                                           #StatConfigDigital[#temp16IndexDigital].OSLevel := #ConfigDint[#temp16IndexDigital].OSLevel;
                                           #StatConfigDigital[#temp16IndexDigital].ApplyExt := #ConfigDint[#temp16IndexDigital].ApplyExt;
                                           #StatConfigDigital[#temp16IndexDigital].ApplyOp := #ConfigDint[#temp16IndexDigital].ApplyOp;
                                           #StatConfigDigital[#temp16IndexDigital].Sync := #ConfigDint[#temp16IndexDigital].Sync;
                                           #StatConfigDigital[#temp16IndexDigital].StateOffOp := #ConfigDint[#temp16IndexDigital].StateOffOp;
                                           #StatConfigDigital[#temp16IndexDigital].StateOpOp := #ConfigDint[#temp16IndexDigital].StateOpOp;
                                           #StatConfigDigital[#temp16IndexDigital].StateAutOp := #ConfigDint[#temp16IndexDigital].StateAutOp;
                                           #StatConfigDigital[#temp16IndexDigital].SrcIntOp := #ConfigDint[#temp16IndexDigital].SrcIntOp;
                                           #StatConfigDigital[#temp16IndexDigital].SrcExtOp := #ConfigDint[#temp16IndexDigital].SrcExtOp;
                                           #StatConfigDigital[#temp16IndexDigital].VExt := #ConfigDint[#temp16IndexDigital].VExt;
                                           #StatConfigDigital[#temp16IndexDigital].VOp := #ConfigDint[#temp16IndexDigital].VOp;
                                       END_IF;
                                       #temp16IndexDigital := #temp16IndexDigital + 1;
                                   END_REGION
                                   // If Parameter type = 3(Binary)
                               #TYPE_BINARY:
                                   REGION Binary
                                       //Bit Masking funtionality for calculate the used Binary parameter
                                       #ConfigParaType.IndexBinary := #ConfigParaType.IndexBinary OR SHL(IN := #temp32TempDword1, N := INT_TO_UINT(#temp16IndexOfDefinition));
                                       //Condition to check the config binary parameters are within range 
                                       IF ((#temp16IndexIO >= #CONFIG_PARAMETER_MIN) AND (#temp16IndexIO <= #MAPPED_CONFIG_BINARY)) THEN
                                           //WinCC Parameter View Faceplate logic
                                           #ConfigBin[#temp16IndexBinary].WQC := #ConfigurationParameterBinary[#temp16IndexMTP].WQC;
                                           #ConfigBin[#temp16IndexBinary].ApplyEn := #ConfigurationParameterBinary[#temp16IndexMTP].ApplyEn;
                                           #ConfigBin[#temp16IndexBinary].ApplyInt := #ConfigurationParameterBinary[#temp16IndexMTP].ApplyInt;
                                           #ConfigBin[#temp16IndexBinary].StateChannel := #ConfigurationParameterBinary[#temp16IndexMTP].StateChannel;
                                           #ConfigBin[#temp16IndexBinary].StateOffAut := #ConfigurationParameterBinary[#temp16IndexMTP].StateOffAut;
                                           #ConfigBin[#temp16IndexBinary].StateOpAut := #ConfigurationParameterBinary[#temp16IndexMTP].StateOpAut;
                                           #ConfigBin[#temp16IndexBinary].StateAutAut := #ConfigurationParameterBinary[#temp16IndexMTP].StateAutAut;
                                           #ConfigBin[#temp16IndexBinary].StateOffAct := #ConfigurationParameterBinary[#temp16IndexMTP].StateOffAct;
                                           #ConfigBin[#temp16IndexBinary].StateOpAct := #ConfigurationParameterBinary[#temp16IndexMTP].StateOpAct;
                                           #ConfigBin[#temp16IndexBinary].StateAutAct := #ConfigurationParameterBinary[#temp16IndexMTP].StateAutAct;
                                           #ConfigBin[#temp16IndexBinary].SrcChannel := #ConfigurationParameterBinary[#temp16IndexMTP].SrcChannel;
                                           #ConfigBin[#temp16IndexBinary].SrcExtAut := #ConfigurationParameterBinary[#temp16IndexMTP].SrcExtAut;
                                           #ConfigBin[#temp16IndexBinary].SrcIntAut := #ConfigurationParameterBinary[#temp16IndexMTP].SrcIntAut;
                                           #ConfigBin[#temp16IndexBinary].SrcIntAct := #ConfigurationParameterBinary[#temp16IndexMTP].SrcIntAct;
                                           #ConfigBin[#temp16IndexBinary].SrcExtAct := #ConfigurationParameterBinary[#temp16IndexMTP].SrcExtAct;
                                           #ConfigBin[#temp16IndexBinary].VInt := #ConfigurationParameterBinary[#temp16IndexMTP].VInt;
                                           #ConfigBin[#temp16IndexBinary].VReq := #ConfigurationParameterBinary[#temp16IndexMTP].VReq;
                                           #ConfigBin[#temp16IndexBinary].VOut := #ConfigurationParameterBinary[#temp16IndexMTP].VOut;
                                           #ConfigBin[#temp16IndexBinary].VFbk := #ConfigurationParameterBinary[#temp16IndexMTP].VFbk;
                                           #ConfigBin[#temp16IndexBinary].VState0 := #ConfigurationParameterBinary[#temp16IndexMTP].VState0;
                                           #ConfigBin[#temp16IndexBinary].VState1 := #ConfigurationParameterBinary[#temp16IndexMTP].VState1;
                                           //Write values from WinCC
                                           IF #ConfigurationParameterBinary[#temp16IndexMTP].OSLevel = #StatConfigBinary[#temp16IndexBinary].OSLevel THEN
                                               #ConfigurationParameterBinary[#temp16IndexMTP].OSLevel := #ConfigBin[#temp16IndexBinary].OSLevel;
                                           ELSE
                                               #ConfigBin[#temp16IndexBinary].OSLevel := #ConfigurationParameterBinary[#temp16IndexMTP].OSLevel;
                                           END_IF;
                                           IF #ConfigurationParameterBinary[#temp16IndexMTP].ApplyExt = #StatConfigBinary[#temp16IndexBinary].ApplyExt THEN
                                               #ConfigurationParameterBinary[#temp16IndexMTP].ApplyExt := #ConfigBin[#temp16IndexBinary].ApplyExt;
                                           ELSE
                                               #ConfigBin[#temp16IndexBinary].ApplyExt := #ConfigurationParameterBinary[#temp16IndexMTP].ApplyExt;
                                           END_IF;
                                           IF #ConfigurationParameterBinary[#temp16IndexMTP].ApplyOp = #StatConfigBinary[#temp16IndexBinary].ApplyOp THEN
                                               #ConfigurationParameterBinary[#temp16IndexMTP].ApplyOp := #ConfigBin[#temp16IndexBinary].ApplyOp;
                                           ELSE
                                               #ConfigBin[#temp16IndexBinary].ApplyOp := #ConfigurationParameterBinary[#temp16IndexMTP].ApplyOp;
                                           END_IF;
                                           IF #ConfigurationParameterBinary[#temp16IndexMTP].Sync = #StatConfigBinary[#temp16IndexBinary].Sync THEN
                                               #ConfigurationParameterBinary[#temp16IndexMTP].Sync := #ConfigBin[#temp16IndexBinary].Sync;
                                           ELSE
                                               #ConfigBin[#temp16IndexBinary].Sync := #ConfigurationParameterBinary[#temp16IndexMTP].Sync;
                                           END_IF;
                                           IF #ConfigurationParameterBinary[#temp16IndexMTP].StateOffOp = #StatConfigBinary[#temp16IndexBinary].StateOffOp THEN
                                               #ConfigurationParameterBinary[#temp16IndexMTP].StateOffOp := #ConfigBin[#temp16IndexBinary].StateOffOp;
                                           ELSE
                                               #ConfigBin[#temp16IndexBinary].StateOffOp := #ConfigurationParameterBinary[#temp16IndexMTP].StateOffOp;
                                           END_IF;
                                           IF #ConfigurationParameterBinary[#temp16IndexMTP].StateOpOp = #StatConfigBinary[#temp16IndexBinary].StateOpOp THEN
                                               #ConfigurationParameterBinary[#temp16IndexMTP].StateOpOp := #ConfigBin[#temp16IndexBinary].StateOpOp;
                                           ELSE
                                               #ConfigBin[#temp16IndexBinary].StateOpOp := #ConfigurationParameterBinary[#temp16IndexMTP].StateOpOp;
                                           END_IF;
                                           IF #ConfigurationParameterBinary[#temp16IndexMTP].StateAutOp = #StatConfigBinary[#temp16IndexBinary].StateAutOp THEN
                                               #ConfigurationParameterBinary[#temp16IndexMTP].StateAutOp := #ConfigBin[#temp16IndexBinary].StateAutOp;
                                           ELSE
                                               #ConfigBin[#temp16IndexBinary].StateAutOp := #ConfigurationParameterBinary[#temp16IndexMTP].StateAutOp;
                                           END_IF;
                                           IF #ConfigurationParameterBinary[#temp16IndexMTP].SrcIntOp = #StatConfigBinary[#temp16IndexBinary].SrcIntOp THEN
                                               #ConfigurationParameterBinary[#temp16IndexMTP].SrcIntOp := #ConfigBin[#temp16IndexBinary].SrcIntOp;
                                           ELSE
                                               #ConfigBin[#temp16IndexBinary].SrcIntOp := #ConfigurationParameterBinary[#temp16IndexMTP].SrcIntOp;
                                           END_IF;
                                           IF #ConfigurationParameterBinary[#temp16IndexMTP].SrcExtOp = #StatConfigBinary[#temp16IndexBinary].SrcExtOp THEN
                                               #ConfigurationParameterBinary[#temp16IndexMTP].SrcExtOp := #ConfigBin[#temp16IndexBinary].SrcExtOp;
                                           ELSE
                                               #ConfigBin[#temp16IndexBinary].SrcExtOp := #ConfigurationParameterBinary[#temp16IndexMTP].SrcExtOp;
                                           END_IF;
                                           IF #ConfigurationParameterBinary[#temp16IndexMTP].VExt = #StatConfigBinary[#temp16IndexBinary].VExt THEN
                                               #ConfigurationParameterBinary[#temp16IndexMTP].VExt := #ConfigBin[#temp16IndexBinary].VExt;
                                           ELSE
                                               #ConfigBin[#temp16IndexBinary].VExt := #ConfigurationParameterBinary[#temp16IndexMTP].VExt;
                                           END_IF;
                                           IF #ConfigurationParameterBinary[#temp16IndexMTP].VOp = #StatConfigBinary[#temp16IndexBinary].VOp THEN
                                               #ConfigurationParameterBinary[#temp16IndexMTP].VOp := #ConfigBin[#temp16IndexBinary].VOp;
                                           ELSE
                                               #ConfigBin[#temp16IndexBinary].VOp := #ConfigurationParameterBinary[#temp16IndexMTP].VOp;
                                           END_IF;

                                           #StatConfigBinary[#temp16IndexBinary].OSLevel := #ConfigBin[#temp16IndexBinary].OSLevel;
                                           #StatConfigBinary[#temp16IndexBinary].ApplyExt := #ConfigBin[#temp16IndexBinary].ApplyExt;
                                           #StatConfigBinary[#temp16IndexBinary].ApplyOp := #ConfigBin[#temp16IndexBinary].ApplyOp;
                                           #StatConfigBinary[#temp16IndexBinary].Sync := #ConfigBin[#temp16IndexBinary].Sync;
                                           #StatConfigBinary[#temp16IndexBinary].StateOffOp := #ConfigBin[#temp16IndexBinary].StateOffOp;
                                           #StatConfigBinary[#temp16IndexBinary].StateOpOp := #ConfigBin[#temp16IndexBinary].StateOpOp;
                                           #StatConfigBinary[#temp16IndexBinary].StateAutOp := #ConfigBin[#temp16IndexBinary].StateAutOp;
                                           #StatConfigBinary[#temp16IndexBinary].SrcIntOp := #ConfigBin[#temp16IndexBinary].SrcIntOp;
                                           #StatConfigBinary[#temp16IndexBinary].SrcExtOp := #ConfigBin[#temp16IndexBinary].SrcExtOp;
                                           #StatConfigBinary[#temp16IndexBinary].VExt := #ConfigBin[#temp16IndexBinary].VExt;
                                           #StatConfigBinary[#temp16IndexBinary].VOp := #ConfigBin[#temp16IndexBinary].VOp;
                                       END_IF;
                                       #temp16IndexBinary := #temp16IndexBinary + 1;
                                   END_REGION
                                   // If Parameter type = 4(String)
                               #TYPE_STRING:
                                   REGION String
                                       //Bit Masking funtionality for calculate the used String parameter
                                       #ConfigParaType.IndexString := #ConfigParaType.IndexString OR SHL(IN := #temp32TempDword1, N := INT_TO_UINT(#temp16IndexOfDefinition));
                                       //Condition to check the config string parameters are within range 
                                       IF ((#temp16IndexIO >= #CONFIG_PARAMETER_MIN) AND (#temp16IndexIO <= #MAPPED_CONFIG_STRING)) THEN
                                           //WinCC Parameter View Faceplate logic
                                           #ConfigString[#temp16IndexString].WQC := #ConfigurationParameterString[#temp16IndexMTP].WQC;
                                           #ConfigString[#temp16IndexString].ApplyEn := #ConfigurationParameterString[#temp16IndexMTP].ApplyEn;
                                           #ConfigString[#temp16IndexString].ApplyInt := #ConfigurationParameterString[#temp16IndexMTP].ApplyInt;
                                           #ConfigString[#temp16IndexString].StateChannel := #ConfigurationParameterString[#temp16IndexMTP].StateChannel;
                                           #ConfigString[#temp16IndexString].StateOffAut := #ConfigurationParameterString[#temp16IndexMTP].StateOffAut;
                                           #ConfigString[#temp16IndexString].StateOpAut := #ConfigurationParameterString[#temp16IndexMTP].StateOpAut;
                                           #ConfigString[#temp16IndexString].StateAutAut := #ConfigurationParameterString[#temp16IndexMTP].StateAutAut;
                                           #ConfigString[#temp16IndexString].StateOffAct := #ConfigurationParameterString[#temp16IndexMTP].StateOffAct;
                                           #ConfigString[#temp16IndexString].StateOpAct := #ConfigurationParameterString[#temp16IndexMTP].StateOpAct;
                                           #ConfigString[#temp16IndexString].StateAutAct := #ConfigurationParameterString[#temp16IndexMTP].StateAutAct;
                                           #ConfigString[#temp16IndexString].SrcChannel := #ConfigurationParameterString[#temp16IndexMTP].SrcChannel;
                                           #ConfigString[#temp16IndexString].SrcExtAut := #ConfigurationParameterString[#temp16IndexMTP].SrcExtAut;
                                           #ConfigString[#temp16IndexString].SrcIntAut := #ConfigurationParameterString[#temp16IndexMTP].SrcIntAut;
                                           #ConfigString[#temp16IndexString].SrcIntAct := #ConfigurationParameterString[#temp16IndexMTP].SrcIntAct;
                                           #ConfigString[#temp16IndexString].SrcExtAct := #ConfigurationParameterString[#temp16IndexMTP].SrcExtAct;
                                           #ConfigString[#temp16IndexString].VInt := #ConfigurationParameterString[#temp16IndexMTP].VInt;
                                           #ConfigString[#temp16IndexString].VReq := #ConfigurationParameterString[#temp16IndexMTP].VReq;
                                           #ConfigString[#temp16IndexString].VOut := #ConfigurationParameterString[#temp16IndexMTP].VOut;
                                           #ConfigString[#temp16IndexString].VFbk := #ConfigurationParameterString[#temp16IndexMTP].VFbk;
                                           //Write values from WinCC
                                           IF #ConfigurationParameterString[#temp16IndexMTP].OSLevel = #StatConfigString[#temp16IndexString].OSLevel THEN
                                               #ConfigurationParameterString[#temp16IndexMTP].OSLevel := #ConfigString[#temp16IndexString].OSLevel;
                                           ELSE
                                               #ConfigString[#temp16IndexString].OSLevel := #ConfigurationParameterString[#temp16IndexMTP].OSLevel;
                                           END_IF;
                                           IF #ConfigurationParameterString[#temp16IndexMTP].ApplyExt = #StatConfigString[#temp16IndexString].ApplyExt THEN
                                               #ConfigurationParameterString[#temp16IndexMTP].ApplyExt := #ConfigString[#temp16IndexString].ApplyExt;
                                           ELSE
                                               #ConfigString[#temp16IndexString].ApplyExt := #ConfigurationParameterString[#temp16IndexMTP].ApplyExt;
                                           END_IF;
                                           IF #ConfigurationParameterString[#temp16IndexMTP].ApplyOp = #StatConfigString[#temp16IndexString].ApplyOp THEN
                                               #ConfigurationParameterString[#temp16IndexMTP].ApplyOp := #ConfigString[#temp16IndexString].ApplyOp;
                                           ELSE
                                               #ConfigString[#temp16IndexString].ApplyOp := #ConfigurationParameterString[#temp16IndexMTP].ApplyOp;
                                           END_IF;
                                           IF #ConfigurationParameterString[#temp16IndexMTP].Sync = #StatConfigString[#temp16IndexString].Sync THEN
                                               #ConfigurationParameterString[#temp16IndexMTP].Sync := #ConfigString[#temp16IndexString].Sync;
                                           ELSE
                                               #ConfigString[#temp16IndexString].Sync := #ConfigurationParameterString[#temp16IndexMTP].Sync;
                                           END_IF;
                                           IF #ConfigurationParameterString[#temp16IndexMTP].StateOffOp = #StatConfigString[#temp16IndexString].StateOffOp THEN
                                               #ConfigurationParameterString[#temp16IndexMTP].StateOffOp := #ConfigString[#temp16IndexString].StateOffOp;
                                           ELSE
                                               #ConfigString[#temp16IndexString].StateOffOp := #ConfigurationParameterString[#temp16IndexMTP].StateOffOp;
                                           END_IF;
                                           IF #ConfigurationParameterString[#temp16IndexMTP].StateOpOp = #StatConfigString[#temp16IndexString].StateOpOp THEN
                                               #ConfigurationParameterString[#temp16IndexMTP].StateOpOp := #ConfigString[#temp16IndexString].StateOpOp;
                                           ELSE
                                               #ConfigString[#temp16IndexString].StateOpOp := #ConfigurationParameterString[#temp16IndexMTP].StateOpOp;
                                           END_IF;
                                           IF #ConfigurationParameterString[#temp16IndexMTP].StateAutOp = #StatConfigString[#temp16IndexString].StateAutOp THEN
                                               #ConfigurationParameterString[#temp16IndexMTP].StateAutOp := #ConfigString[#temp16IndexString].StateAutOp;
                                           ELSE
                                               #ConfigString[#temp16IndexString].StateAutOp := #ConfigurationParameterString[#temp16IndexMTP].StateAutOp;
                                           END_IF;
                                           IF #ConfigurationParameterString[#temp16IndexMTP].SrcIntOp = #StatConfigString[#temp16IndexString].SrcIntOp THEN
                                               #ConfigurationParameterString[#temp16IndexMTP].SrcIntOp := #ConfigString[#temp16IndexString].SrcIntOp;
                                           ELSE
                                               #ConfigString[#temp16IndexString].SrcIntOp := #ConfigurationParameterString[#temp16IndexMTP].SrcIntOp;
                                           END_IF;
                                           IF #ConfigurationParameterString[#temp16IndexMTP].SrcExtOp = #StatConfigString[#temp16IndexString].SrcExtOp THEN
                                               #ConfigurationParameterString[#temp16IndexMTP].SrcExtOp := #ConfigString[#temp16IndexString].SrcExtOp;
                                           ELSE
                                               #ConfigString[#temp16IndexString].SrcExtOp := #ConfigurationParameterString[#temp16IndexMTP].SrcExtOp;
                                           END_IF;
                                           IF #ConfigurationParameterString[#temp16IndexMTP].VExt = #StatConfigString[#temp16IndexString].VExt THEN
                                               #ConfigurationParameterString[#temp16IndexMTP].VExt := #ConfigString[#temp16IndexString].VExt;
                                           ELSE
                                               #ConfigString[#temp16IndexString].VExt := #ConfigurationParameterString[#temp16IndexMTP].VExt;
                                           END_IF;
                                           IF #ConfigurationParameterString[#temp16IndexMTP].VOp = #StatConfigString[#temp16IndexString].VOp THEN
                                               #ConfigurationParameterString[#temp16IndexMTP].VOp := #ConfigString[#temp16IndexString].VOp;
                                           ELSE
                                               #ConfigString[#temp16IndexString].VOp := #ConfigurationParameterString[#temp16IndexMTP].VOp;
                                           END_IF;

                                           #StatConfigString[#temp16IndexString].OSLevel := #ConfigString[#temp16IndexString].OSLevel;
                                           #StatConfigString[#temp16IndexString].ApplyExt := #ConfigString[#temp16IndexString].ApplyExt;
                                           #StatConfigString[#temp16IndexString].ApplyOp := #ConfigString[#temp16IndexString].ApplyOp;
                                           #StatConfigString[#temp16IndexString].Sync := #ConfigString[#temp16IndexString].Sync;
                                           #StatConfigString[#temp16IndexString].StateOffOp := #ConfigString[#temp16IndexString].StateOffOp;
                                           #StatConfigString[#temp16IndexString].StateOpOp := #ConfigString[#temp16IndexString].StateOpOp;
                                           #StatConfigString[#temp16IndexString].StateAutOp := #ConfigString[#temp16IndexString].StateAutOp;
                                           #StatConfigString[#temp16IndexString].SrcIntOp := #ConfigString[#temp16IndexString].SrcIntOp;
                                           #StatConfigString[#temp16IndexString].SrcExtOp := #ConfigString[#temp16IndexString].SrcExtOp;
                                           #StatConfigString[#temp16IndexString].VExt := #ConfigString[#temp16IndexString].VExt;
                                           #StatConfigString[#temp16IndexString].VOp := #ConfigString[#temp16IndexString].VOp;
                                       END_IF;
                                       #temp16IndexString := #temp16IndexString + 1;
                                   END_REGION
                           END_CASE;
                       END_IF;
                   END_IF;
               END_FOR;
           END_IF;
       END_REGION
      REGION Procedure Parameter
           REGION Get Current/Prepared procedure ID
               //Get Current procedure index number from setup DB
               IF (#ProcedureCur > 0) THEN
                   FOR #temp16i := #NUMBER_OF_PROCEDURES_MIN TO #NUMBER_OF_PROCEDURES BY 1 DO
                       IF #ProcedureCur = #tempSetup.procedure.procedure[#temp16i].Procedure.ProcedureID THEN
                           #stat16ProceCurIndex := #temp16i;
                           EXIT;
                       END_IF;
                   END_FOR;
               END_IF;
               //Get Prepared procedure index number from setup DB
               IF (#ProcedureReq> 0) THEN
                   FOR #temp16i := #NUMBER_OF_PROCEDURES_MIN TO #NUMBER_OF_PROCEDURES BY 1 DO
                       IF #ProcedureReq = #tempSetup.procedure.procedure[#temp16i].Procedure.ProcedureID THEN
                           #stat16ProceReqIndex := #temp16i;
                           EXIT;
                       END_IF;
                   END_FOR;
               END_IF;
           END_REGION
           REGION Get Start and End index details of the Current /Prepared procedure
               //Current/Prepared procedure selection for parameter display in the faceplate
               IF NOT (#ProcedureParaType.ProcedureReqCurInd) THEN
                   //Get current Procedure step order details from Starting State
                   #tempProcStartingStartIndex := #tempSetup.procedure.procedure[#stat16ProceCurIndex].StateTransient.starting.startIndex;
                   #tempProcStartingEndIndex := #tempSetup.procedure.procedure[#stat16ProceCurIndex].StateTransient.starting.endIndex;
                   //Get current Procedure step order details from Running State
                   #tempProcRunningStartIndex := #tempSetup.procedure.procedure[#stat16ProceCurIndex].StateTransient.running.startIndex;
                   #tempProcRunningEndIndex := #tempSetup.procedure.procedure[#stat16ProceCurIndex].StateTransient.running.endIndex;
                   //Get current Procedure step order details from Holding State
                   #tempProcHoldingStartIndex := #tempSetup.procedure.procedure[#stat16ProceCurIndex].StateTransient.holding.startIndex;
                   #tempProcHoldingEndIndex := #tempSetup.procedure.procedure[#stat16ProceCurIndex].StateTransient.holding.endIndex;
                   //Get current Procedure step order details from unholding State
                   #tempProcUnHoldingStartIndex := #tempSetup.procedure.procedure[#stat16ProceCurIndex].StateTransient.unholding.startIndex;
                   #tempProcUnHoldingEndIndex := #tempSetup.procedure.procedure[#stat16ProceCurIndex].StateTransient.unholding.endIndex;
                   //Get current Procedure step order details from pausing State
                   #tempProcUnPausingStartIndex := #tempSetup.procedure.procedure[#stat16ProceCurIndex].StateTransient.pausing.startIndex;
                   #tempProcUnPausingEndIndex := #tempSetup.procedure.procedure[#stat16ProceCurIndex].StateTransient.pausing.endIndex;
                   //Get current Procedure step order details from resuming State
                   #tempProcResumingStartIndex := #tempSetup.procedure.procedure[#stat16ProceCurIndex].StateTransient.resuming.startIndex;
                   #tempProcResumingEndIndex := #tempSetup.procedure.procedure[#stat16ProceCurIndex].StateTransient.resuming.endIndex;
                   //Get current Procedure step order details from completing State
                   #tempProcCompletingStartIndex := #tempSetup.procedure.procedure[#stat16ProceCurIndex].StateTransient.completing.startIndex;
                   #tempProcCompletingEndIndex := #tempSetup.procedure.procedure[#stat16ProceCurIndex].StateTransient.completing.endIndex;
                   //Get current Procedure step order details from stopping State
                   #tempProcStoppingStartIndex := #tempSetup.procedure.procedure[#stat16ProceCurIndex].StateTransient.stopping.startIndex;
                   #tempProcStoppingEndIndex := #tempSetup.procedure.procedure[#stat16ProceCurIndex].StateTransient.stopping.endIndex;
                   //Get current Procedure step order details from aborting State
                   #tempProcAbortingStartIndex := #tempSetup.procedure.procedure[#stat16ProceCurIndex].StateTransient.aborting.startIndex;
                   #tempProcAbortingEndIndex := #tempSetup.procedure.procedure[#stat16ProceCurIndex].StateTransient.aborting.endIndex;
                   //Get current Procedure step order details from resetting State
                   #tempProcResettingStartIndex := #tempSetup.procedure.procedure[#stat16ProceCurIndex].StateTransient.resetting.startIndex;
                   #tempProcResettingEndIndex := #tempSetup.procedure.procedure[#stat16ProceCurIndex].StateTransient.resetting.endIndex;

               ELSIF (#ProcedureParaType.ProcedureReqCurInd) THEN
                   //Get current Procedure step order details from Starting State
                   #tempProcStartingStartIndex := #tempSetup.procedure.procedure[#stat16ProceReqIndex].StateTransient.starting.startIndex;
                   #tempProcStartingEndIndex := #tempSetup.procedure.procedure[#stat16ProceReqIndex].StateTransient.starting.endIndex;
                   //Get current Procedure step order details from Running State
                   #tempProcRunningStartIndex := #tempSetup.procedure.procedure[#stat16ProceReqIndex].StateTransient.running.startIndex;
                   #tempProcRunningEndIndex := #tempSetup.procedure.procedure[#stat16ProceReqIndex].StateTransient.running.endIndex;
                   //Get current Procedure step order details from Holding State
                   #tempProcHoldingStartIndex := #tempSetup.procedure.procedure[#stat16ProceReqIndex].StateTransient.holding.startIndex;
                   #tempProcHoldingEndIndex := #tempSetup.procedure.procedure[#stat16ProceReqIndex].StateTransient.holding.endIndex;
                   //Get current Procedure step order details from unholding State
                   #tempProcUnHoldingStartIndex := #tempSetup.procedure.procedure[#stat16ProceReqIndex].StateTransient.unholding.startIndex;
                   #tempProcUnHoldingEndIndex := #tempSetup.procedure.procedure[#stat16ProceReqIndex].StateTransient.unholding.endIndex;
                   //Get current Procedure step order details from pausing State
                   #tempProcUnPausingStartIndex := #tempSetup.procedure.procedure[#stat16ProceReqIndex].StateTransient.pausing.startIndex;
                   #tempProcUnPausingEndIndex := #tempSetup.procedure.procedure[#stat16ProceReqIndex].StateTransient.pausing.endIndex;
                   //Get current Procedure step order details from resuming State
                   #tempProcResumingStartIndex := #tempSetup.procedure.procedure[#stat16ProceReqIndex].StateTransient.resuming.startIndex;
                   #tempProcResumingEndIndex := #tempSetup.procedure.procedure[#stat16ProceReqIndex].StateTransient.resuming.endIndex;
                   //Get current Procedure step order details from completing State
                   #tempProcCompletingStartIndex := #tempSetup.procedure.procedure[#stat16ProceReqIndex].StateTransient.completing.startIndex;
                   #tempProcCompletingEndIndex := #tempSetup.procedure.procedure[#stat16ProceReqIndex].StateTransient.completing.endIndex;
                   //Get current Procedure step order details from stopping State
                   #tempProcStoppingStartIndex := #tempSetup.procedure.procedure[#stat16ProceReqIndex].StateTransient.stopping.startIndex;
                   #tempProcStoppingEndIndex := #tempSetup.procedure.procedure[#stat16ProceReqIndex].StateTransient.stopping.endIndex;
                   //Get current Procedure step order details from aborting State
                   #tempProcAbortingStartIndex := #tempSetup.procedure.procedure[#stat16ProceReqIndex].StateTransient.aborting.startIndex;
                   #tempProcAbortingEndIndex := #tempSetup.procedure.procedure[#stat16ProceReqIndex].StateTransient.aborting.endIndex;
                   //Get current Procedure step order details from resetting State
                   #tempProcResettingStartIndex := #tempSetup.procedure.procedure[#stat16ProceReqIndex].StateTransient.resetting.startIndex;
                   #tempProcResettingEndIndex := #tempSetup.procedure.procedure[#stat16ProceReqIndex].StateTransient.resetting.endIndex;
               END_IF;

               #tempProcStartIndex := -1;
               #tempProcEndIndex := -1;
               //Get the Start and End index from the States
               IF (#tempProcStartingStartIndex > -1) AND (#tempProcStartingEndIndex > -1) THEN
                   #tempProcStartIndex := #tempProcStartingStartIndex;
                   #tempProcEndIndex := #tempProcStartingEndIndex;
               ELSIF (#tempProcRunningStartIndex > -1) AND (#tempProcRunningEndIndex > -1) THEN
                   #tempProcStartIndex := #tempProcRunningStartIndex;
                   #tempProcEndIndex := #tempProcRunningEndIndex;
               ELSIF (#tempProcHoldingStartIndex > -1) AND (#tempProcHoldingEndIndex > -1) THEN
                   #tempProcStartIndex := #tempProcHoldingStartIndex;
                   #tempProcEndIndex := #tempProcHoldingEndIndex;
               ELSIF (#tempProcUnHoldingStartIndex > -1) AND (#tempProcUnHoldingEndIndex > -1) THEN
                   #tempProcStartIndex := #tempProcUnHoldingStartIndex;
                   #tempProcEndIndex := #tempProcUnHoldingEndIndex;
               ELSIF (#tempProcUnPausingStartIndex > -1) AND (#tempProcUnPausingEndIndex > -1) THEN
                   #tempProcStartIndex := #tempProcUnPausingStartIndex;
                   #tempProcEndIndex := #tempProcUnPausingEndIndex;
               ELSIF (#tempProcResumingStartIndex > -1) AND (#tempProcResumingEndIndex > -1) THEN
                   #tempProcStartIndex := #tempProcResumingStartIndex;
                   #tempProcEndIndex := #tempProcResumingEndIndex;
               ELSIF (#tempProcCompletingStartIndex > -1) AND (#tempProcCompletingEndIndex > -1) THEN
                   #tempProcStartIndex := #tempProcCompletingStartIndex;
                   #tempProcEndIndex := #tempProcCompletingEndIndex;
               ELSIF (#tempProcStoppingStartIndex > -1) AND (#tempProcStoppingEndIndex > -1) THEN
                   #tempProcStartIndex := #tempProcStoppingStartIndex;
                   #tempProcEndIndex := #tempProcStoppingEndIndex;
               ELSIF (#tempProcAbortingStartIndex > -1) AND (#tempProcAbortingEndIndex > -1) THEN
                   #tempProcStartIndex := #tempProcAbortingStartIndex;
                   #tempProcEndIndex := #tempProcAbortingEndIndex;
               ELSIF (#tempProcResettingStartIndex > -1) AND (#tempProcResettingEndIndex > -1) THEN
                   #tempProcStartIndex := #tempProcResettingStartIndex;
                   #tempProcEndIndex := #tempProcResettingEndIndex;
               END_IF;

               //Get Current Procedure step order parameter index details
               IF (#tempProcStartIndex > -1) AND (#tempProcEndIndex > -1) THEN
                   #stat16ProcParaStartIndex := #tempSetup.stepOrder.stepOrder[#tempProcStartIndex].parameter.startIndex;
                   #stat16ProcParaEndIndex := #tempSetup.stepOrder.stepOrder[#tempProcEndIndex].parameter.endIndex;
               END_IF;
           END_REGION


           REGION Get mapped/used procedure parameters and move to the procedure parameter FP variables
               // Condition to check the start and end index values is within the range
               IF ((#stat16ProcParaStartIndex >= #PARAMETERINDEX_MIN) AND (#stat16ProcParaStartIndex <= #PARAMETERINDEX_MAX))
                   AND ((#stat16ProcParaEndIndex >= #PARAMETERINDEX_MIN) AND (#stat16ProcParaEndIndex <= #PARAMETERINDEX_MAX))
                   AND ((#stat16ProcParaEndIndex - #stat16ProcParaStartIndex + #PROCEDURE_PARAMETER_MIN) <= #PROCEDURE_PARAMETER_MAX) THEN

                   //Initialize the used variable values
                   #temp32TempDword1 := 16#1;
                   #temp16IndexAnalog := 16#0;
                   #temp16IndexDigital := 16#0;
                   #temp16IndexBinary := 16#0;
                   #temp16IndexString := 16#0;
                   //Initialize the Procedure Para index and Name index while changing of Procedure and changing of screen selection b/w Prepared and Current procedure
                   IF ((#statLasProcedureCur <> #ProcedureCur) OR (#statLasProcedureReq <> #ProcedureReq) OR (#statLastReqProcedSelected <> #ProcedureParaType.ProcedureReqCurInd)) THEN
                       #ProcedureParaType.IndexAnalog := 16#0;
                       #ProcedureParaType.NameIndexAnalog := 16#0;
                       #ProcedureParaType.IndexDigital := 16#0;
                       #ProcedureParaType.NameIndexDigital := 16#0;
                       #ProcedureParaType.IndexBinary := 16#0;
                       #ProcedureParaType.NameIndexBinary := 16#0;
                       #ProcedureParaType.IndexString := 16#0;
                       #ProcedureParaType.NameIndexString := 16#0;
                   END_IF;
                   IF (((#ProcedureCur <> 16#0) AND NOT #ProcedureParaType.ProcedureReqCurInd) OR ((#ProcedureReq <> 16#0) AND #ProcedureParaType.ProcedureReqCurInd)) THEN
                       //Used/Mapped parameter count with individual parameter type will written from the Tool
                       #statTotalProcedureParameters := #MAPPED_PROCEDURE_ANALOG + #MAPPED_PROCEDURE_DIGITAL + #MAPPED_PROCEDURE_BINARY + #MAPPED_PROCEDURE_STRING - 1;
                       IF ((#statTotalProcedureParameters >= 0) AND (#statTotalProcedureParameters <= #PROCEDURE_PARAMETER_MAX)) THEN
                           FOR #temp16IndexOfDefinition := #PROCEDURE_PARAMETER_MIN TO #statTotalProcedureParameters BY 1 DO
                               // Condition for allow the loop iteration only within the start and end index
                               IF (((#stat16ProcParaEndIndex - #stat16ProcParaStartIndex) - #temp16IndexOfDefinition + #PROCEDURE_PARAMETER_MIN) >= 0) THEN
                                   #statInternalCurProcParameter[#temp16IndexOfDefinition].index := #tempSetup.stepOrder.parameterIndex[#stat16ProcParaStartIndex + #temp16IndexOfDefinition];  // MiS: content of first parameterIndex to first internal index, content of second parameterIndex to second internal index etc.
                                   #temp16Index := #statInternalCurProcParameter[#temp16IndexOfDefinition].index;//Move index info to the local var
                                   #temp16ParameterType := #tempSetup.step.parameterDefinition[#temp16Index].type;  // Get type of current parameter
                                   #temp16IndexMTP := #tempSetup.step.parameterDefinition[#temp16Index].indexMTP;//Get parameter indexMTP(wrapper DB) from the setup DB.
                                   #temp16IndexIO := #tempSetup.step.parameterDefinition[#temp16Index].indexIO;
                                   //Condition TO check parameter types are in the range
                                   IF (#temp16ParameterType >= #TYPE_NONE) AND (#temp16ParameterType <= #TYPE_STRING) THEN
                                       REGION Copy procedure parameters from input
                                           CASE #temp16ParameterType OF
                                                   // If Parameter type = 1(Analog)
                                               #TYPE_ANALOG:
                                                   REGION Analog
                                                       //Bit Masking funtionality for calculate the used Analog parameter and Position of the Parameter name in the HMI Text List                                              
                                                       #ProcedureParaType.IndexAnalog := #ProcedureParaType.IndexAnalog OR SHL(IN := #temp32TempDword1, N := INT_TO_UINT(#temp16IndexOfDefinition));
                                                       #ProcedureParaType.NameIndexAnalog := #ProcedureParaType.NameIndexAnalog OR SHL(IN := #temp32TempDword1, N := INT_TO_UINT(#temp16Index));
                                                       //WinCC Parameter View Faceplate logic
                                                       //#StatConfigPara.Analog[#temp16IndexIO] := #MTPConfigurationParameterAnalog[#temp16IndexMTP];
                                                       #ProcedureAna[#temp16IndexAnalog].WQC := #ProcedureParameterAnalog[#temp16IndexMTP].WQC;
                                                       #ProcedureAna[#temp16IndexAnalog].ApplyEn := #ProcedureParameterAnalog[#temp16IndexMTP].ApplyEn;
                                                       #ProcedureAna[#temp16IndexAnalog].ApplyInt := #ProcedureParameterAnalog[#temp16IndexMTP].ApplyInt;
                                                       #ProcedureAna[#temp16IndexAnalog].StateChannel := #ProcedureParameterAnalog[#temp16IndexMTP].StateChannel;
                                                       #ProcedureAna[#temp16IndexAnalog].StateOffAut := #ProcedureParameterAnalog[#temp16IndexMTP].StateOffAut;
                                                       #ProcedureAna[#temp16IndexAnalog].StateOpAut := #ProcedureParameterAnalog[#temp16IndexMTP].StateOpAut;
                                                       #ProcedureAna[#temp16IndexAnalog].StateAutAut := #ProcedureParameterAnalog[#temp16IndexMTP].StateAutAut;
                                                       #ProcedureAna[#temp16IndexAnalog].StateOffAct := #ProcedureParameterAnalog[#temp16IndexMTP].StateOffAct;
                                                       #ProcedureAna[#temp16IndexAnalog].StateOpAct := #ProcedureParameterAnalog[#temp16IndexMTP].StateOpAct;
                                                       #ProcedureAna[#temp16IndexAnalog].StateAutAct := #ProcedureParameterAnalog[#temp16IndexMTP].StateAutAct;
                                                       #ProcedureAna[#temp16IndexAnalog].SrcChannel := #ProcedureParameterAnalog[#temp16IndexMTP].SrcChannel;
                                                       #ProcedureAna[#temp16IndexAnalog].SrcExtAut := #ProcedureParameterAnalog[#temp16IndexMTP].SrcExtAut;
                                                       #ProcedureAna[#temp16IndexAnalog].SrcIntAut := #ProcedureParameterAnalog[#temp16IndexMTP].SrcIntAut;
                                                       #ProcedureAna[#temp16IndexAnalog].SrcIntAct := #ProcedureParameterAnalog[#temp16IndexMTP].SrcIntAct;
                                                       #ProcedureAna[#temp16IndexAnalog].SrcExtAct := #ProcedureParameterAnalog[#temp16IndexMTP].SrcExtAct;
                                                       #ProcedureAna[#temp16IndexAnalog].VInt := #ProcedureParameterAnalog[#temp16IndexMTP].VInt;
                                                       #ProcedureAna[#temp16IndexAnalog].VReq := #ProcedureParameterAnalog[#temp16IndexMTP].VReq;
                                                       #ProcedureAna[#temp16IndexAnalog].VOut := #ProcedureParameterAnalog[#temp16IndexMTP].VOut;
                                                       #ProcedureAna[#temp16IndexAnalog].VFbk := #ProcedureParameterAnalog[#temp16IndexMTP].VFbk;
                                                       #ProcedureAna[#temp16IndexAnalog].VSclMin := #ProcedureParameterAnalog[#temp16IndexMTP].VSclMin;
                                                       #ProcedureAna[#temp16IndexAnalog].VSclMax := #ProcedureParameterAnalog[#temp16IndexMTP].VSclMax;
                                                       #ProcedureAna[#temp16IndexAnalog].VUnit := #ProcedureParameterAnalog[#temp16IndexMTP].VUnit;
                                                       #ProcedureAna[#temp16IndexAnalog].VMin := #ProcedureParameterAnalog[#temp16IndexMTP].VMin;
                                                       #ProcedureAna[#temp16IndexAnalog].VMax := #ProcedureParameterAnalog[#temp16IndexMTP].VMax;
                                                       //Write values from WinCC
                                                       IF #ProcedureParameterAnalog[#temp16IndexMTP].OSLevel = #StatProcedureAnalog[#temp16IndexAnalog].OSLevel THEN
                                                           #ProcedureParameterAnalog[#temp16IndexMTP].OSLevel := #ProcedureAna[#temp16IndexAnalog].OSLevel;
                                                       ELSE
                                                           #ProcedureAna[#temp16IndexAnalog].OSLevel := #ProcedureParameterAnalog[#temp16IndexMTP].OSLevel;
                                                       END_IF;
                                                       IF #ProcedureParameterAnalog[#temp16IndexMTP].ApplyExt = #StatProcedureAnalog[#temp16IndexAnalog].ApplyExt THEN
                                                           #ProcedureParameterAnalog[#temp16IndexMTP].ApplyExt := #ProcedureAna[#temp16IndexAnalog].ApplyExt;
                                                       ELSE
                                                           #ProcedureAna[#temp16IndexAnalog].ApplyExt := #ProcedureParameterAnalog[#temp16IndexMTP].ApplyExt;
                                                       END_IF;
                                                       IF #ProcedureParameterAnalog[#temp16IndexMTP].ApplyOp = #StatProcedureAnalog[#temp16IndexAnalog].ApplyOp THEN
                                                           #ProcedureParameterAnalog[#temp16IndexMTP].ApplyOp := #ProcedureAna[#temp16IndexAnalog].ApplyOp;
                                                       ELSE
                                                           #ProcedureAna[#temp16IndexAnalog].ApplyOp := #ProcedureParameterAnalog[#temp16IndexMTP].ApplyOp;
                                                       END_IF;
                                                       IF #ProcedureParameterAnalog[#temp16IndexMTP].Sync = #StatProcedureAnalog[#temp16IndexAnalog].Sync THEN
                                                           #ProcedureParameterAnalog[#temp16IndexMTP].Sync := #ProcedureAna[#temp16IndexAnalog].Sync;
                                                       ELSE
                                                           #ProcedureAna[#temp16IndexAnalog].Sync := #ProcedureParameterAnalog[#temp16IndexMTP].Sync;
                                                       END_IF;
                                                       IF #ProcedureParameterAnalog[#temp16IndexMTP].StateOffOp = #StatProcedureAnalog[#temp16IndexAnalog].StateOffOp THEN
                                                           #ProcedureParameterAnalog[#temp16IndexMTP].StateOffOp := #ProcedureAna[#temp16IndexAnalog].StateOffOp;
                                                       ELSE
                                                           #ProcedureAna[#temp16IndexAnalog].StateOffOp := #ProcedureParameterAnalog[#temp16IndexMTP].StateOffOp;
                                                       END_IF;
                                                       IF #ProcedureParameterAnalog[#temp16IndexMTP].StateOpOp = #StatProcedureAnalog[#temp16IndexAnalog].StateOpOp THEN
                                                           #ProcedureParameterAnalog[#temp16IndexMTP].StateOpOp := #ProcedureAna[#temp16IndexAnalog].StateOpOp;
                                                       ELSE
                                                           #ProcedureAna[#temp16IndexAnalog].StateOpOp := #ProcedureParameterAnalog[#temp16IndexMTP].StateOpOp;
                                                       END_IF;
                                                       IF #ProcedureParameterAnalog[#temp16IndexMTP].StateAutOp = #StatProcedureAnalog[#temp16IndexAnalog].StateAutOp THEN
                                                           #ProcedureParameterAnalog[#temp16IndexMTP].StateAutOp := #ProcedureAna[#temp16IndexAnalog].StateAutOp;
                                                       ELSE
                                                           #ProcedureAna[#temp16IndexAnalog].StateAutOp := #ProcedureParameterAnalog[#temp16IndexMTP].StateAutOp;
                                                       END_IF;
                                                       IF #ProcedureParameterAnalog[#temp16IndexMTP].SrcIntOp = #StatProcedureAnalog[#temp16IndexAnalog].SrcIntOp THEN
                                                           #ProcedureParameterAnalog[#temp16IndexMTP].SrcIntOp := #ProcedureAna[#temp16IndexAnalog].SrcIntOp;
                                                       ELSE
                                                           #ProcedureAna[#temp16IndexAnalog].SrcIntOp := #ProcedureParameterAnalog[#temp16IndexMTP].SrcIntOp;
                                                       END_IF;
                                                       IF #ProcedureParameterAnalog[#temp16IndexMTP].SrcExtOp = #StatProcedureAnalog[#temp16IndexAnalog].SrcExtOp THEN
                                                           #ProcedureParameterAnalog[#temp16IndexMTP].SrcExtOp := #ProcedureAna[#temp16IndexAnalog].SrcExtOp;
                                                       ELSE
                                                           #ProcedureAna[#temp16IndexAnalog].SrcExtOp := #ProcedureParameterAnalog[#temp16IndexMTP].SrcExtOp;
                                                       END_IF;
                                                       IF #ProcedureParameterAnalog[#temp16IndexMTP].VExt = #StatProcedureAnalog[#temp16IndexAnalog].VExt THEN
                                                           #ProcedureParameterAnalog[#temp16IndexMTP].VExt := #ProcedureAna[#temp16IndexAnalog].VExt;
                                                       ELSE
                                                           #ProcedureAna[#temp16IndexAnalog].VExt := #ProcedureParameterAnalog[#temp16IndexMTP].VExt;
                                                       END_IF;
                                                       IF #ProcedureParameterAnalog[#temp16IndexMTP].VOp = #StatProcedureAnalog[#temp16IndexAnalog].VOp THEN
                                                           #ProcedureParameterAnalog[#temp16IndexMTP].VOp := #ProcedureAna[#temp16IndexAnalog].VOp;
                                                       ELSE
                                                           #ProcedureAna[#temp16IndexAnalog].VOp := #ProcedureParameterAnalog[#temp16IndexMTP].VOp;
                                                       END_IF;

                                                       #StatProcedureAnalog[#temp16IndexAnalog].OSLevel := #ProcedureAna[#temp16IndexAnalog].OSLevel;
                                                       #StatProcedureAnalog[#temp16IndexAnalog].ApplyExt := #ProcedureAna[#temp16IndexAnalog].ApplyExt;
                                                       #StatProcedureAnalog[#temp16IndexAnalog].ApplyOp := #ProcedureAna[#temp16IndexAnalog].ApplyOp;
                                                       #StatProcedureAnalog[#temp16IndexAnalog].Sync := #ProcedureAna[#temp16IndexAnalog].Sync;
                                                       #StatProcedureAnalog[#temp16IndexAnalog].StateOffOp := #ProcedureAna[#temp16IndexAnalog].StateOffOp;
                                                       #StatProcedureAnalog[#temp16IndexAnalog].StateOpOp := #ProcedureAna[#temp16IndexAnalog].StateOpOp;
                                                       #StatProcedureAnalog[#temp16IndexAnalog].StateAutOp := #ProcedureAna[#temp16IndexAnalog].StateAutOp;
                                                       #StatProcedureAnalog[#temp16IndexAnalog].SrcIntOp := #ProcedureAna[#temp16IndexAnalog].SrcIntOp;
                                                       #StatProcedureAnalog[#temp16IndexAnalog].SrcExtOp := #ProcedureAna[#temp16IndexAnalog].SrcExtOp;
                                                       #StatProcedureAnalog[#temp16IndexAnalog].VExt := #ProcedureAna[#temp16IndexAnalog].VExt;
                                                       #StatProcedureAnalog[#temp16IndexAnalog].VOp := #ProcedureAna[#temp16IndexAnalog].VOp;

                                                       #temp16IndexAnalog := #temp16IndexAnalog + 1;
                                                   END_REGION
                                                   // If Parameter type = 2(Digital)     
                                               #TYPE_DIGITAL:
                                                   REGION Digital
                                                       //Bit Masking funtionality for calculate the used Digital parameter and Position of the Parameter name in the HMI Text List  
                                                       #ProcedureParaType.IndexDigital := #ProcedureParaType.IndexDigital OR SHL(IN := #temp32TempDword1, N := INT_TO_UINT(#temp16IndexOfDefinition));
                                                       #ProcedureParaType.NameIndexDigital := #ProcedureParaType.NameIndexDigital OR SHL(IN := #temp32TempDword1, N := INT_TO_UINT(#temp16Index));
                                                       //WinCC Parameter View Faceplate logic
                                                       //#StatConfigPara.Digital[#temp16IndexIO] := #MTPConfigurationParameterAnalog[#temp16IndexMTP];
                                                       #ProcedureDint[#temp16IndexDigital].WQC := #ProcedureParameterDigital[#temp16IndexMTP].WQC;
                                                       #ProcedureDint[#temp16IndexDigital].ApplyEn := #ProcedureParameterDigital[#temp16IndexMTP].ApplyEn;
                                                       #ProcedureDint[#temp16IndexDigital].ApplyInt := #ProcedureParameterDigital[#temp16IndexMTP].ApplyInt;
                                                       #ProcedureDint[#temp16IndexDigital].StateChannel := #ProcedureParameterDigital[#temp16IndexMTP].StateChannel;
                                                       #ProcedureDint[#temp16IndexDigital].StateOffAut := #ProcedureParameterDigital[#temp16IndexMTP].StateOffAut;
                                                       #ProcedureDint[#temp16IndexDigital].StateOpAut := #ProcedureParameterDigital[#temp16IndexMTP].StateOpAut;
                                                       #ProcedureDint[#temp16IndexDigital].StateAutAut := #ProcedureParameterDigital[#temp16IndexMTP].StateAutAut;
                                                       #ProcedureDint[#temp16IndexDigital].StateOffAct := #ProcedureParameterDigital[#temp16IndexMTP].StateOffAct;
                                                       #ProcedureDint[#temp16IndexDigital].StateOpAct := #ProcedureParameterDigital[#temp16IndexMTP].StateOpAct;
                                                       #ProcedureDint[#temp16IndexDigital].StateAutAct := #ProcedureParameterDigital[#temp16IndexMTP].StateAutAct;
                                                       #ProcedureDint[#temp16IndexDigital].SrcChannel := #ProcedureParameterDigital[#temp16IndexMTP].SrcChannel;
                                                       #ProcedureDint[#temp16IndexDigital].SrcExtAut := #ProcedureParameterDigital[#temp16IndexMTP].SrcExtAut;
                                                       #ProcedureDint[#temp16IndexDigital].SrcIntAut := #ProcedureParameterDigital[#temp16IndexMTP].SrcIntAut;
                                                       #ProcedureDint[#temp16IndexDigital].SrcIntAct := #ProcedureParameterDigital[#temp16IndexMTP].SrcIntAct;
                                                       #ProcedureDint[#temp16IndexDigital].SrcExtAct := #ProcedureParameterDigital[#temp16IndexMTP].SrcExtAct;
                                                       #ProcedureDint[#temp16IndexDigital].VInt := #ProcedureParameterDigital[#temp16IndexMTP].VInt;
                                                       #ProcedureDint[#temp16IndexDigital].VReq := #ProcedureParameterDigital[#temp16IndexMTP].VReq;
                                                       #ProcedureDint[#temp16IndexDigital].VOut := #ProcedureParameterDigital[#temp16IndexMTP].VOut;
                                                       #ProcedureDint[#temp16IndexDigital].VFbk := #ProcedureParameterDigital[#temp16IndexMTP].VFbk;
                                                       #ProcedureDint[#temp16IndexDigital].VSclMin := #ProcedureParameterDigital[#temp16IndexMTP].VSclMin;
                                                       #ProcedureDint[#temp16IndexDigital].VSclMax := #ProcedureParameterDigital[#temp16IndexMTP].VSclMax;
                                                       #ProcedureDint[#temp16IndexDigital].VUnit := #ProcedureParameterDigital[#temp16IndexMTP].VUnit;
                                                       #ProcedureDint[#temp16IndexDigital].VMin := #ProcedureParameterDigital[#temp16IndexMTP].VMin;
                                                       #ProcedureDint[#temp16IndexDigital].VMax := #ProcedureParameterDigital[#temp16IndexMTP].VMax;
                                                       //Write values from WinCC
                                                       IF #ProcedureParameterDigital[#temp16IndexMTP].OSLevel = #StatProcedureDigital[#temp16IndexDigital].OSLevel THEN
                                                           #ProcedureParameterDigital[#temp16IndexMTP].OSLevel := #ProcedureDint[#temp16IndexDigital].OSLevel;
                                                       ELSE
                                                           #ProcedureDint[#temp16IndexDigital].OSLevel := #ProcedureParameterDigital[#temp16IndexMTP].OSLevel;
                                                       END_IF;
                                                       IF #ProcedureParameterDigital[#temp16IndexMTP].ApplyExt = #StatProcedureDigital[#temp16IndexDigital].ApplyExt THEN
                                                           #ProcedureParameterDigital[#temp16IndexMTP].ApplyExt := #ProcedureDint[#temp16IndexDigital].ApplyExt;
                                                       ELSE
                                                           #ProcedureDint[#temp16IndexDigital].ApplyExt := #ProcedureParameterDigital[#temp16IndexMTP].ApplyExt;
                                                       END_IF;
                                                       IF #ProcedureParameterDigital[#temp16IndexMTP].ApplyOp = #StatProcedureDigital[#temp16IndexDigital].ApplyOp THEN
                                                           #ProcedureParameterDigital[#temp16IndexMTP].ApplyOp := #ProcedureDint[#temp16IndexDigital].ApplyOp;
                                                       ELSE
                                                           #ProcedureDint[#temp16IndexDigital].ApplyOp := #ProcedureParameterDigital[#temp16IndexMTP].ApplyOp;
                                                       END_IF;
                                                       IF #ProcedureParameterDigital[#temp16IndexMTP].Sync = #StatProcedureDigital[#temp16IndexDigital].Sync THEN
                                                           #ProcedureParameterDigital[#temp16IndexMTP].Sync := #ProcedureDint[#temp16IndexDigital].Sync;
                                                       ELSE
                                                           #ProcedureDint[#temp16IndexDigital].Sync := #ProcedureParameterDigital[#temp16IndexMTP].Sync;
                                                       END_IF;
                                                       IF #ProcedureParameterDigital[#temp16IndexMTP].StateOffOp = #StatProcedureDigital[#temp16IndexDigital].StateOffOp THEN
                                                           #ProcedureParameterDigital[#temp16IndexMTP].StateOffOp := #ProcedureDint[#temp16IndexDigital].StateOffOp;
                                                       ELSE
                                                           #ProcedureDint[#temp16IndexDigital].StateOffOp := #ProcedureParameterDigital[#temp16IndexMTP].StateOffOp;
                                                       END_IF;
                                                       IF #ProcedureParameterDigital[#temp16IndexMTP].StateOpOp = #StatProcedureDigital[#temp16IndexDigital].StateOpOp THEN
                                                           #ProcedureParameterDigital[#temp16IndexMTP].StateOpOp := #ProcedureDint[#temp16IndexDigital].StateOpOp;
                                                       ELSE
                                                           #ProcedureDint[#temp16IndexDigital].StateOpOp := #ProcedureParameterDigital[#temp16IndexMTP].StateOpOp;
                                                       END_IF;
                                                       IF #ProcedureParameterDigital[#temp16IndexMTP].StateAutOp = #StatProcedureDigital[#temp16IndexDigital].StateAutOp THEN
                                                           #ProcedureParameterDigital[#temp16IndexMTP].StateAutOp := #ProcedureDint[#temp16IndexDigital].StateAutOp;
                                                       ELSE
                                                           #ProcedureDint[#temp16IndexDigital].StateAutOp := #ProcedureParameterDigital[#temp16IndexMTP].StateAutOp;
                                                       END_IF;
                                                       IF #ProcedureParameterDigital[#temp16IndexMTP].SrcIntOp = #StatProcedureDigital[#temp16IndexDigital].SrcIntOp THEN
                                                           #ProcedureParameterDigital[#temp16IndexMTP].SrcIntOp := #ProcedureDint[#temp16IndexDigital].SrcIntOp;
                                                       ELSE
                                                           #ProcedureDint[#temp16IndexDigital].SrcIntOp := #ProcedureParameterDigital[#temp16IndexMTP].SrcIntOp;
                                                       END_IF;
                                                       IF #ProcedureParameterDigital[#temp16IndexMTP].SrcExtOp = #StatProcedureDigital[#temp16IndexDigital].SrcExtOp THEN
                                                           #ProcedureParameterDigital[#temp16IndexMTP].SrcExtOp := #ProcedureDint[#temp16IndexDigital].SrcExtOp;
                                                       ELSE
                                                           #ProcedureDint[#temp16IndexDigital].SrcExtOp := #ProcedureParameterDigital[#temp16IndexMTP].SrcExtOp;
                                                       END_IF;
                                                       IF #ProcedureParameterDigital[#temp16IndexMTP].VExt = #StatProcedureDigital[#temp16IndexDigital].VExt THEN
                                                           #ProcedureParameterDigital[#temp16IndexMTP].VExt := #ProcedureDint[#temp16IndexDigital].VExt;
                                                       ELSE
                                                           #ProcedureDint[#temp16IndexDigital].VExt := #ProcedureParameterDigital[#temp16IndexMTP].VExt;
                                                       END_IF;
                                                       IF #ProcedureParameterDigital[#temp16IndexMTP].VOp = #StatProcedureDigital[#temp16IndexDigital].VOp THEN
                                                           #ProcedureParameterDigital[#temp16IndexMTP].VOp := #ProcedureDint[#temp16IndexDigital].VOp;
                                                       ELSE
                                                           #ProcedureDint[#temp16IndexDigital].VOp := #ProcedureParameterDigital[#temp16IndexMTP].VOp;
                                                       END_IF;

                                                       #StatProcedureDigital[#temp16IndexDigital].OSLevel := #ProcedureDint[#temp16IndexDigital].OSLevel;
                                                       #StatProcedureDigital[#temp16IndexDigital].ApplyExt := #ProcedureDint[#temp16IndexDigital].ApplyExt;
                                                       #StatProcedureDigital[#temp16IndexDigital].ApplyOp := #ProcedureDint[#temp16IndexDigital].ApplyOp;
                                                       #StatProcedureDigital[#temp16IndexDigital].Sync := #ProcedureDint[#temp16IndexDigital].Sync;
                                                       #StatProcedureDigital[#temp16IndexDigital].StateOffOp := #ProcedureDint[#temp16IndexDigital].StateOffOp;
                                                       #StatProcedureDigital[#temp16IndexDigital].StateOpOp := #ProcedureDint[#temp16IndexDigital].StateOpOp;
                                                       #StatProcedureDigital[#temp16IndexDigital].StateAutOp := #ProcedureDint[#temp16IndexDigital].StateAutOp;
                                                       #StatProcedureDigital[#temp16IndexDigital].SrcIntOp := #ProcedureDint[#temp16IndexDigital].SrcIntOp;
                                                       #StatProcedureDigital[#temp16IndexDigital].SrcExtOp := #ProcedureDint[#temp16IndexDigital].SrcExtOp;
                                                       #StatProcedureDigital[#temp16IndexDigital].VExt := #ProcedureDint[#temp16IndexDigital].VExt;
                                                       #StatProcedureDigital[#temp16IndexDigital].VOp := #ProcedureDint[#temp16IndexDigital].VOp;

                                                       #temp16IndexDigital := #temp16IndexDigital + 1;
                                                   END_REGION
                                                   // If Parameter type = 3(Binary)    
                                               #TYPE_BINARY:
                                                   REGION Binary
                                                       //Bit Masking funtionality for calculate the used Binary parameter and Position of the Parameter name in the HMI Text List  
                                                       #ProcedureParaType.IndexBinary := #ProcedureParaType.IndexBinary OR SHL(IN := #temp32TempDword1, N := INT_TO_UINT(#temp16IndexOfDefinition));
                                                       #ProcedureParaType.NameIndexBinary := #ProcedureParaType.NameIndexBinary OR SHL(IN := #temp32TempDword1, N := INT_TO_UINT(#temp16Index));
                                                       //WinCC Parameter View Faceplate logic
                                                       //#StatConfigPara.Binary[#temp16IndexIO] := #MTPConfigurationParameterAnalog[#temp16IndexMTP];
                                                       #ProcedureBin[#temp16IndexBinary].WQC := #ProcedureParameterBinary[#temp16IndexMTP].WQC;
                                                       #ProcedureBin[#temp16IndexBinary].ApplyEn := #ProcedureParameterBinary[#temp16IndexMTP].ApplyEn;
                                                       #ProcedureBin[#temp16IndexBinary].ApplyInt := #ProcedureParameterBinary[#temp16IndexMTP].ApplyInt;
                                                       #ProcedureBin[#temp16IndexBinary].StateChannel := #ProcedureParameterBinary[#temp16IndexMTP].StateChannel;
                                                       #ProcedureBin[#temp16IndexBinary].StateOffAut := #ProcedureParameterBinary[#temp16IndexMTP].StateOffAut;
                                                       #ProcedureBin[#temp16IndexBinary].StateOpAut := #ProcedureParameterBinary[#temp16IndexMTP].StateOpAut;
                                                       #ProcedureBin[#temp16IndexBinary].StateAutAut := #ProcedureParameterBinary[#temp16IndexMTP].StateAutAut;
                                                       #ProcedureBin[#temp16IndexBinary].StateOffAct := #ProcedureParameterBinary[#temp16IndexMTP].StateOffAct;
                                                       #ProcedureBin[#temp16IndexBinary].StateOpAct := #ProcedureParameterBinary[#temp16IndexMTP].StateOpAct;
                                                       #ProcedureBin[#temp16IndexBinary].StateAutAct := #ProcedureParameterBinary[#temp16IndexMTP].StateAutAct;
                                                       #ProcedureBin[#temp16IndexBinary].SrcChannel := #ProcedureParameterBinary[#temp16IndexMTP].SrcChannel;
                                                       #ProcedureBin[#temp16IndexBinary].SrcExtAut := #ProcedureParameterBinary[#temp16IndexMTP].SrcExtAut;
                                                       #ProcedureBin[#temp16IndexBinary].SrcIntAut := #ProcedureParameterBinary[#temp16IndexMTP].SrcIntAut;
                                                       #ProcedureBin[#temp16IndexBinary].SrcIntAct := #ProcedureParameterBinary[#temp16IndexMTP].SrcIntAct;
                                                       #ProcedureBin[#temp16IndexBinary].SrcExtAct := #ProcedureParameterBinary[#temp16IndexMTP].SrcExtAct;
                                                       #ProcedureBin[#temp16IndexBinary].VInt := #ProcedureParameterBinary[#temp16IndexMTP].VInt;
                                                       #ProcedureBin[#temp16IndexBinary].VReq := #ProcedureParameterBinary[#temp16IndexMTP].VReq;
                                                       #ProcedureBin[#temp16IndexBinary].VOut := #ProcedureParameterBinary[#temp16IndexMTP].VOut;
                                                       #ProcedureBin[#temp16IndexBinary].VFbk := #ProcedureParameterBinary[#temp16IndexMTP].VFbk;

                                                       //Write values from WinCC
                                                       IF #ProcedureParameterBinary[#temp16IndexMTP].OSLevel = #StatProcedureBinary[#temp16IndexBinary].OSLevel THEN
                                                           #ProcedureParameterBinary[#temp16IndexMTP].OSLevel := #ProcedureBin[#temp16IndexBinary].OSLevel;
                                                       ELSE
                                                           #ProcedureBin[#temp16IndexBinary].OSLevel := #ProcedureParameterBinary[#temp16IndexMTP].OSLevel;
                                                       END_IF;
                                                       IF #ProcedureParameterBinary[#temp16IndexMTP].ApplyExt = #StatProcedureBinary[#temp16IndexBinary].ApplyExt THEN
                                                           #ProcedureParameterBinary[#temp16IndexMTP].ApplyExt := #ProcedureBin[#temp16IndexBinary].ApplyExt;
                                                       ELSE
                                                           #ProcedureBin[#temp16IndexBinary].ApplyExt := #ProcedureParameterBinary[#temp16IndexMTP].ApplyExt;
                                                       END_IF;
                                                       IF #ProcedureParameterBinary[#temp16IndexMTP].ApplyOp = #StatProcedureBinary[#temp16IndexBinary].ApplyOp THEN
                                                           #ProcedureParameterBinary[#temp16IndexMTP].ApplyOp := #ProcedureBin[#temp16IndexBinary].ApplyOp;
                                                       ELSE
                                                           #ProcedureBin[#temp16IndexBinary].ApplyOp := #ProcedureParameterBinary[#temp16IndexMTP].ApplyOp;
                                                       END_IF;
                                                       IF #ProcedureParameterBinary[#temp16IndexMTP].Sync = #StatProcedureBinary[#temp16IndexBinary].Sync THEN
                                                           #ProcedureParameterBinary[#temp16IndexMTP].Sync := #ProcedureBin[#temp16IndexBinary].Sync;
                                                       ELSE
                                                           #ProcedureBin[#temp16IndexBinary].Sync := #ProcedureParameterBinary[#temp16IndexMTP].Sync;
                                                       END_IF;
                                                       IF #ProcedureParameterBinary[#temp16IndexMTP].StateOffOp = #StatProcedureBinary[#temp16IndexBinary].StateOffOp THEN
                                                           #ProcedureParameterBinary[#temp16IndexMTP].StateOffOp := #ProcedureBin[#temp16IndexBinary].StateOffOp;
                                                       ELSE
                                                           #ProcedureBin[#temp16IndexBinary].StateOffOp := #ProcedureParameterBinary[#temp16IndexMTP].StateOffOp;
                                                       END_IF;
                                                       IF #ProcedureParameterBinary[#temp16IndexMTP].StateOpOp = #StatProcedureBinary[#temp16IndexBinary].StateOpOp THEN
                                                           #ProcedureParameterBinary[#temp16IndexMTP].StateOpOp := #ProcedureBin[#temp16IndexBinary].StateOpOp;
                                                       ELSE
                                                           #ProcedureBin[#temp16IndexBinary].StateOpOp := #ProcedureParameterBinary[#temp16IndexMTP].StateOpOp;
                                                       END_IF;
                                                       IF #ProcedureParameterBinary[#temp16IndexMTP].StateAutOp = #StatProcedureBinary[#temp16IndexBinary].StateAutOp THEN
                                                           #ProcedureParameterBinary[#temp16IndexMTP].StateAutOp := #ProcedureBin[#temp16IndexBinary].StateAutOp;
                                                       ELSE
                                                           #ProcedureBin[#temp16IndexBinary].StateAutOp := #ProcedureParameterBinary[#temp16IndexMTP].StateAutOp;
                                                       END_IF;
                                                       IF #ProcedureParameterBinary[#temp16IndexMTP].SrcIntOp = #StatProcedureBinary[#temp16IndexBinary].SrcIntOp THEN
                                                           #ProcedureParameterBinary[#temp16IndexMTP].SrcIntOp := #ProcedureBin[#temp16IndexBinary].SrcIntOp;
                                                       ELSE
                                                           #ProcedureBin[#temp16IndexBinary].SrcIntOp := #ProcedureParameterBinary[#temp16IndexMTP].SrcIntOp;
                                                       END_IF;
                                                       IF #ProcedureParameterBinary[#temp16IndexMTP].SrcExtOp = #StatProcedureBinary[#temp16IndexBinary].SrcExtOp THEN
                                                           #ProcedureParameterBinary[#temp16IndexMTP].SrcExtOp := #ProcedureBin[#temp16IndexBinary].SrcExtOp;
                                                       ELSE
                                                           #ProcedureBin[#temp16IndexBinary].SrcExtOp := #ProcedureParameterBinary[#temp16IndexMTP].SrcExtOp;
                                                       END_IF;
                                                       IF #ProcedureParameterBinary[#temp16IndexMTP].VExt = #StatProcedureBinary[#temp16IndexBinary].VExt THEN
                                                           #ProcedureParameterBinary[#temp16IndexMTP].VExt := #ProcedureBin[#temp16IndexBinary].VExt;
                                                       ELSE
                                                           #ProcedureBin[#temp16IndexBinary].VExt := #ProcedureParameterBinary[#temp16IndexMTP].VExt;
                                                       END_IF;
                                                       IF #ProcedureParameterBinary[#temp16IndexMTP].VOp = #StatProcedureBinary[#temp16IndexBinary].VOp THEN
                                                           #ProcedureParameterBinary[#temp16IndexMTP].VOp := #ProcedureBin[#temp16IndexBinary].VOp;
                                                       ELSE
                                                           #ProcedureBin[#temp16IndexBinary].VOp := #ProcedureParameterBinary[#temp16IndexMTP].VOp;
                                                       END_IF;

                                                       #StatProcedureBinary[#temp16IndexBinary].OSLevel := #ProcedureBin[#temp16IndexBinary].OSLevel;
                                                       #StatProcedureBinary[#temp16IndexBinary].ApplyExt := #ProcedureBin[#temp16IndexBinary].ApplyExt;
                                                       #StatProcedureBinary[#temp16IndexBinary].ApplyOp := #ProcedureBin[#temp16IndexBinary].ApplyOp;
                                                       #StatProcedureBinary[#temp16IndexBinary].Sync := #ProcedureBin[#temp16IndexBinary].Sync;
                                                       #StatProcedureBinary[#temp16IndexBinary].StateOffOp := #ProcedureBin[#temp16IndexBinary].StateOffOp;
                                                       #StatProcedureBinary[#temp16IndexBinary].StateOpOp := #ProcedureBin[#temp16IndexBinary].StateOpOp;
                                                       #StatProcedureBinary[#temp16IndexBinary].StateAutOp := #ProcedureBin[#temp16IndexBinary].StateAutOp;
                                                       #StatProcedureBinary[#temp16IndexBinary].SrcIntOp := #ProcedureBin[#temp16IndexBinary].SrcIntOp;
                                                       #StatProcedureBinary[#temp16IndexBinary].SrcExtOp := #ProcedureBin[#temp16IndexBinary].SrcExtOp;
                                                       #StatProcedureBinary[#temp16IndexBinary].VExt := #ProcedureBin[#temp16IndexBinary].VExt;
                                                       #StatProcedureBinary[#temp16IndexBinary].VOp := #ProcedureBin[#temp16IndexBinary].VOp;

                                                       #temp16IndexBinary := #temp16IndexBinary + 1;
                                                   END_REGION
                                                   // If Parameter type = 4(String)    
                                               #TYPE_STRING:
                                                   REGION String
                                                       //Bit Masking funtionality for calculate the used String parameter and Position of the Parameter name in the HMI Text List  
                                                       #ProcedureParaType.IndexString := #ProcedureParaType.IndexString OR SHL(IN := #temp32TempDword1, N := INT_TO_UINT(#temp16IndexOfDefinition));
                                                       #ProcedureParaType.NameIndexString := #ProcedureParaType.NameIndexString OR SHL(IN := #temp32TempDword1, N := INT_TO_UINT(#temp16Index));
                                                       //WinCC Parameter View Faceplate logic
                                                       //#StatConfigPara."String"[#temp16IndexIO] := #MTPConfigurationParameterString[#temp16IndexMTP];
                                                       #ProcedureString[#temp16IndexString].WQC := #ProcedureParameterString[#temp16IndexMTP].WQC;
                                                       #ProcedureString[#temp16IndexString].ApplyEn := #ProcedureParameterString[#temp16IndexMTP].ApplyEn;
                                                       #ProcedureString[#temp16IndexString].ApplyInt := #ProcedureParameterString[#temp16IndexMTP].ApplyInt;
                                                       #ProcedureString[#temp16IndexString].StateChannel := #ProcedureParameterString[#temp16IndexMTP].StateChannel;
                                                       #ProcedureString[#temp16IndexString].StateOffAut := #ProcedureParameterString[#temp16IndexMTP].StateOffAut;
                                                       #ProcedureString[#temp16IndexString].StateOpAut := #ProcedureParameterString[#temp16IndexMTP].StateOpAut;
                                                       #ProcedureString[#temp16IndexString].StateAutAut := #ProcedureParameterString[#temp16IndexMTP].StateAutAut;
                                                       #ProcedureString[#temp16IndexString].StateOffAct := #ProcedureParameterString[#temp16IndexMTP].StateOffAct;
                                                       #ProcedureString[#temp16IndexString].StateOpAct := #ProcedureParameterString[#temp16IndexMTP].StateOpAct;
                                                       #ProcedureString[#temp16IndexString].StateAutAct := #ProcedureParameterString[#temp16IndexMTP].StateAutAct;
                                                       #ProcedureString[#temp16IndexString].SrcChannel := #ProcedureParameterString[#temp16IndexMTP].SrcChannel;
                                                       #ProcedureString[#temp16IndexString].SrcExtAut := #ProcedureParameterString[#temp16IndexMTP].SrcExtAut;
                                                       #ProcedureString[#temp16IndexString].SrcIntAut := #ProcedureParameterString[#temp16IndexMTP].SrcIntAut;
                                                       #ProcedureString[#temp16IndexString].SrcIntAct := #ProcedureParameterString[#temp16IndexMTP].SrcIntAct;
                                                       #ProcedureString[#temp16IndexString].SrcExtAct := #ProcedureParameterString[#temp16IndexMTP].SrcExtAct;
                                                       #ProcedureString[#temp16IndexString].VInt := #ProcedureParameterString[#temp16IndexMTP].VInt;
                                                       #ProcedureString[#temp16IndexString].VReq := #ProcedureParameterString[#temp16IndexMTP].VReq;
                                                       #ProcedureString[#temp16IndexString].VOut := #ProcedureParameterString[#temp16IndexMTP].VOut;
                                                       #ProcedureString[#temp16IndexString].VFbk := #ProcedureParameterString[#temp16IndexMTP].VFbk;

                                                       //Write values from WinCC
                                                       IF #ProcedureParameterString[#temp16IndexMTP].OSLevel = #StatProcedureString[#temp16IndexString].OSLevel THEN
                                                           #ProcedureParameterString[#temp16IndexMTP].OSLevel := #ProcedureString[#temp16IndexString].OSLevel;
                                                       ELSE
                                                           #ProcedureString[#temp16IndexString].OSLevel := #ProcedureParameterString[#temp16IndexMTP].OSLevel;
                                                       END_IF;
                                                       IF #ProcedureParameterString[#temp16IndexMTP].ApplyExt = #StatProcedureString[#temp16IndexString].ApplyExt THEN
                                                           #ProcedureParameterString[#temp16IndexMTP].ApplyExt := #ProcedureString[#temp16IndexString].ApplyExt;
                                                       ELSE
                                                           #ProcedureString[#temp16IndexString].ApplyExt := #ProcedureParameterString[#temp16IndexMTP].ApplyExt;
                                                       END_IF;
                                                       IF #ProcedureParameterString[#temp16IndexMTP].ApplyOp = #StatProcedureString[#temp16IndexString].ApplyOp THEN
                                                           #ProcedureParameterString[#temp16IndexMTP].ApplyOp := #ProcedureString[#temp16IndexString].ApplyOp;
                                                       ELSE
                                                           #ProcedureString[#temp16IndexString].ApplyOp := #ProcedureParameterString[#temp16IndexMTP].ApplyOp;
                                                       END_IF;
                                                       IF #ProcedureParameterString[#temp16IndexMTP].Sync = #StatProcedureString[#temp16IndexString].Sync THEN
                                                           #ProcedureParameterString[#temp16IndexMTP].Sync := #ProcedureString[#temp16IndexString].Sync;
                                                       ELSE
                                                           #ProcedureString[#temp16IndexString].Sync := #ProcedureParameterString[#temp16IndexMTP].Sync;
                                                       END_IF;
                                                       IF #ProcedureParameterString[#temp16IndexMTP].StateOffOp = #StatProcedureString[#temp16IndexString].StateOffOp THEN
                                                           #ProcedureParameterString[#temp16IndexMTP].StateOffOp := #ProcedureString[#temp16IndexString].StateOffOp;
                                                       ELSE
                                                           #ProcedureString[#temp16IndexString].StateOffOp := #ProcedureParameterString[#temp16IndexMTP].StateOffOp;
                                                       END_IF;
                                                       IF #ProcedureParameterString[#temp16IndexMTP].StateOpOp = #StatProcedureString[#temp16IndexString].StateOpOp THEN
                                                           #ProcedureParameterString[#temp16IndexMTP].StateOpOp := #ProcedureString[#temp16IndexString].StateOpOp;
                                                       ELSE
                                                           #ProcedureString[#temp16IndexString].StateOpOp := #ProcedureParameterString[#temp16IndexMTP].StateOpOp;
                                                       END_IF;
                                                       IF #ProcedureParameterString[#temp16IndexMTP].StateAutOp = #StatProcedureString[#temp16IndexString].StateAutOp THEN
                                                           #ProcedureParameterString[#temp16IndexMTP].StateAutOp := #ProcedureString[#temp16IndexString].StateAutOp;
                                                       ELSE
                                                           #ProcedureString[#temp16IndexString].StateAutOp := #ProcedureParameterString[#temp16IndexMTP].StateAutOp;
                                                       END_IF;
                                                       IF #ProcedureParameterString[#temp16IndexMTP].SrcIntOp = #StatProcedureString[#temp16IndexString].SrcIntOp THEN
                                                           #ProcedureParameterString[#temp16IndexMTP].SrcIntOp := #ProcedureString[#temp16IndexString].SrcIntOp;
                                                       ELSE
                                                           #ProcedureString[#temp16IndexString].SrcIntOp := #ProcedureParameterString[#temp16IndexMTP].SrcIntOp;
                                                       END_IF;
                                                       IF #ProcedureParameterString[#temp16IndexMTP].SrcExtOp = #StatProcedureString[#temp16IndexString].SrcExtOp THEN
                                                           #ProcedureParameterString[#temp16IndexMTP].SrcExtOp := #ProcedureString[#temp16IndexString].SrcExtOp;
                                                       ELSE
                                                           #ProcedureString[#temp16IndexString].SrcExtOp := #ProcedureParameterString[#temp16IndexMTP].SrcExtOp;
                                                       END_IF;
                                                       IF #ProcedureParameterString[#temp16IndexMTP].VExt = #StatProcedureString[#temp16IndexString].VExt THEN
                                                           #ProcedureParameterString[#temp16IndexMTP].VExt := #ProcedureString[#temp16IndexString].VExt;
                                                       ELSE
                                                           #ProcedureString[#temp16IndexString].VExt := #ProcedureParameterString[#temp16IndexMTP].VExt;
                                                       END_IF;
                                                       IF #ProcedureParameterString[#temp16IndexMTP].VOp = #StatProcedureString[#temp16IndexString].VOp THEN
                                                           #ProcedureParameterString[#temp16IndexMTP].VOp := #ProcedureString[#temp16IndexString].VOp;
                                                       ELSE
                                                           #ProcedureString[#temp16IndexString].VOp := #ProcedureParameterString[#temp16IndexMTP].VOp;
                                                       END_IF;

                                                       #StatProcedureString[#temp16IndexString].OSLevel := #ProcedureString[#temp16IndexString].OSLevel;
                                                       #StatProcedureString[#temp16IndexString].ApplyExt := #ProcedureString[#temp16IndexString].ApplyExt;
                                                       #StatProcedureString[#temp16IndexString].ApplyOp := #ProcedureString[#temp16IndexString].ApplyOp;
                                                       #StatProcedureString[#temp16IndexString].Sync := #ProcedureString[#temp16IndexString].Sync;
                                                       #StatProcedureString[#temp16IndexString].StateOffOp := #ProcedureString[#temp16IndexString].StateOffOp;
                                                       #StatProcedureString[#temp16IndexString].StateOpOp := #ProcedureString[#temp16IndexString].StateOpOp;
                                                       #StatProcedureString[#temp16IndexString].StateAutOp := #ProcedureString[#temp16IndexString].StateAutOp;
                                                       #StatProcedureString[#temp16IndexString].SrcIntOp := #ProcedureString[#temp16IndexString].SrcIntOp;
                                                       #StatProcedureString[#temp16IndexString].SrcExtOp := #ProcedureString[#temp16IndexString].SrcExtOp;
                                                       #StatProcedureString[#temp16IndexString].VExt := #ProcedureString[#temp16IndexString].VExt;
                                                       #StatProcedureString[#temp16IndexString].VOp := #ProcedureString[#temp16IndexString].VOp;

                                                       #temp16IndexString := #temp16IndexString + 1;
                                                   END_REGION
                                           END_CASE;
                                       END_REGION
                                   END_IF;
                               END_IF;
                           END_FOR;
                       END_IF;
                   END_IF;
               END_IF;
           END_REGION
       END_REGION

       REGION Process In Values

           REGION Get Start and End index details of the Current /Prepared procedure
               //Current/Prepared procedure selection for parameter display in the faceplate
               //#stat32PrecedureProcessInMap := -1;
               IF NOT (#ProcessInValueType.ProcedureReqCurInd) THEN
                   #stat32PrecedureProcessInMap := #tempSetup.procedure.procedure[#stat16ProceCurIndex].ProcedureProcessInMap[0];
               ELSIF (#ProcessInValueType.ProcedureReqCurInd) THEN
                   #stat32PrecedureProcessInMap := #tempSetup.procedure.procedure[#stat16ProceReqIndex].ProcedureProcessInMap[0];
               END_IF;
           END_REGION
           //Initialize the used variable values        
           #temp32TempDword1 := 16#1;
           #temp16IndexAnalog := 16#0;
           #temp16IndexDigital := 16#0;
           #temp16IndexBinary := 16#0;
           #temp16IndexString := 16#0;
           //Initialize the Process In Value index and Name index while changing of Procedure and changing of screen selection b/w Prepared and Current procedure
           IF ((#statLasProcedureCur <> #ProcedureCur) OR (#statLasProcedureReq <> #ProcedureReq) OR (#StatLastProceselProcessIn <> #ProcessInValueType.ProcedureReqCurInd)
               OR (((#ProcedureCur = 16#0) AND NOT #ProcessInValueType.ProcedureReqCurInd) OR ((#ProcedureReq = 16#0) AND #ProcessInValueType.ProcedureReqCurInd))) THEN
               #ProcessInValueType.IndexAnalog := 16#0;
               #ProcessInValueType.NameIndexAnalog := 16#0;
               #ProcessInValueType.IndexDigital := 16#0;
               #ProcessInValueType.NameIndexDigital := 16#0;
               #ProcessInValueType.IndexBinary := 16#0;
               #ProcessInValueType.NameIndexBinary := 16#0;
               #ProcessInValueType.IndexString := 16#0;
               #ProcessInValueType.NameIndexString := 16#0;
           END_IF;
           //Used/Mapped parameter count with individual parameter type will written from the Tool
           #statTotalProcessInValues := #MAPPED_PROCESS_IN_ANALOG + #MAPPED_PROCESS_IN_DIGITAL + #MAPPED_PROCESS_IN_BINARY + #MAPPED_PROCESS_IN_STRING - 1;
           IF (((#ProcedureCur <> 16#0) AND NOT #ProcessInValueType.ProcedureReqCurInd) OR ((#ProcedureReq <> 16#0) AND #ProcessInValueType.ProcedureReqCurInd)) THEN
               IF ((#statTotalProcessInValues >= 0) AND (#statTotalProcessInValues <= #PROCESS_VALUES_IN_MAX)) THEN
                   #temp16IndexOfDefinitionProcessIn := 16#0;
                   FOR #temp16IndexOfDefinition := #PROCESS_VALUES_IN_MIN TO #statTotalProcessInValues BY 1 DO
                       #temp16ParameterCMAddress := BYTE_TO_INT(#tempSetup.processValueInData.definition[#temp16IndexOfDefinition].controlModule);
                       #temp16ParameterType := #tempSetup.processValueInData.definition[#temp16IndexOfDefinition].type;
                       #temp16IndexMTP := #tempSetup.processValueInData.definition[#temp16IndexOfDefinition].indexMTP;
                       #tempUsed := #tempSetup.processValueInData.used;
                       // Find the procedure information assigned with the processIn values
                       IF (((#stat32PrecedureProcessInMap AND SHL(IN := #temp32TempDword1, N := INT_TO_UINT(#temp16IndexOfDefinition))) <> 0) = TRUE) THEN
                           #temp16IndexIO := #tempSetup.processValueInData.definition[#temp16IndexOfDefinition].indexIO;

